Fanuc KAREL source: compact_preamble.KL

PROGRAM KB00026
%NOLOCKGROUP
%ENVIRONMENT REGOPE
VAR
P1:INTEGER;P2:INTEGER;P3:INTEGER
BEGIN
P1=1
P2=1
P3=1
CLR_POS_REG(P1,P2,P3)
END KB00026
